FUNCTION F_CtrlIn: LREAL
(*
Function used to set input of controller.

Constructor: 		Patryk Panylo
Company:		E. Riexinger GmbH
Date:			03.06.2014
Version:			1.00

Date:			Revision:		Who:				Comment
dd.mm.yyyy		x.xx			Initials			comment

*)
VAR_INPUT
	(* Enummerations *)

	(* Variables *)
	lrSetPoint							:LREAL;							(* Set point - SP *)
	lrProcessVariable						:LREAL;							(* Process variable - PV *)
	lrDeadZone							:LREAL;							(* Dead zone - noise*)

	(* References *)

	(* Interfaces *)

	(* Instances *)

END_VAR
VAR
END_VAR


F_CtrlIn := F_DeadZone(
	lrSetPoint - lrProcessVariable,
	lrDeadZone
);

END_FUNCTION

(* stored: Version 1.1.0.1, ProductVersion 3.1.4024.15
   POU F_CtrlIn: Id {6a177f74-27ed-4834-942c-c19208b1cc2b}, SpecialFunc None *)
